Fanuc KAREL source: kt00238.KL

-- PROVISIONAL review KL for V1013-1; original PC SHA256 b3ce4d0a6411afe9cec305ff68afcc7b233fef20bccfaa8e704de79eab879623
-- Incomplete behavior may be omitted. Consult companion uncertainty JSON. Do not deploy.
PROGRAM KT00238
%NOLOCKGROUP
VAR
  I1 : INTEGER
  OUT : INTEGER
-- UNRESOLVED_DECL Y2 type=002018
BEGIN
  -- UNRESOLVED_PC offsets 5-16; opcodes 2E,23
  -- UNRESOLVED_PC offsets 21-35; opcodes 2E,22,9D,33,B2
  -- UNRESOLVED_PC offsets 40-62; opcodes 21,22,9D,33,B1,47,23
  -- UNRESOLVED_PC offsets 67-71; opcodes 7F
END KT00238
